RoboDK station: POC(1).rdk

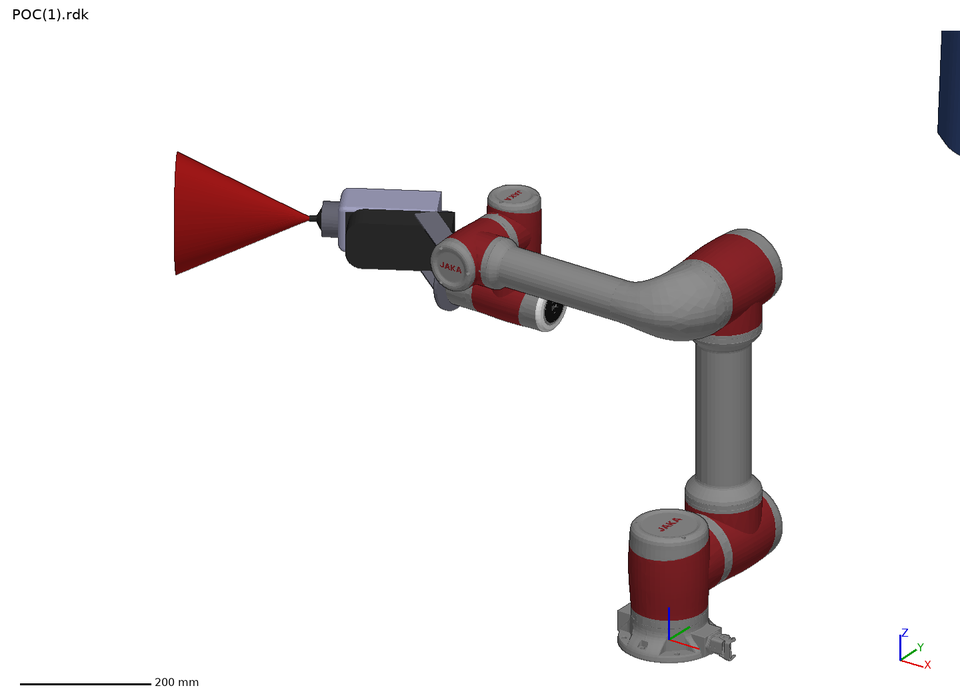
[picture v0: the station drawn from its stored meshes, robots at their saved joint values, targets as dots, program paths as lines]
Station POC(1) (saved by RoboDK 6.2.2). Poses are relative to the parent item; angles as X-Y-Z fixed-axis rotations.
  - frame JAKA Zu5 Base at (0, 0, 0) mm
    - robot JAKA Zu5: 6 axes, payload 5 kg, reach 954 mm, repeatability 0.02 mm, weight 23 kg
        modified DH rows (alpha deg, a mm, theta deg, d mm): 0, 0, 0, 120.15; 90, 0, 0, 0; 0, 430, 0, 0; 0, 368.5, -180, -114; -90, 0, 0, 113.5; 90, 0, 180, 107
        joint limits [-360, -85, -175, -85, -360, -360] to [360, 265, 175, 265, 360, 360]; home [0, 90, 90, 180, 90, 0]; saved at [0, 90, 90, 180, 90, 0]
      - tool Paint gun, TCP at (50, 0, 450) mm, rotated rx 0 ry 30 rz 0 deg, size 203.2 x 279.7 x 471.5 mm
  - object Denim_Surface at (0, 0, 0) mm, size 353.8 x 49.4 x 413.5 mm
